// Résultats d'une action (docs/04 § 5)
{attribute 'pack_mode' := '1'}
TYPE ST_ActResults :
STRUCT
    nCount : USINT;
    aReal : ARRAY[1..GVL_Const.MAX_PARAMS] OF LREAL;
    aJudgement : ARRAY[1..GVL_Const.MAX_PARAMS] OF E_Judgement;
    stPos : ST_Position;        // le résultat de type Position, s'il y en a un
    nPosIndex : USINT;          // rang du résultat de type Position, 0 = aucun
    sText : STRING(80);         // le résultat de type Text, s'il y en a un
    nTextIndex : USINT;         // rang du résultat de type Text, 0 = aucun
END_STRUCT
END_TYPE

(* stored: Version 1.1.0.1, ProductVersion 3.1.4024.12
   DUT ST_ActResults: Id {a5f5fd08-d8d5-56b6-81e8-6d68d7fcfb8e} *)
